// TIA Portal V21 export
DATA_BLOCK "Issue221_unitNested_readOnly"   // DB
{ S7_Optimized_Access := 'TRUE' }
// stored: AutoNumber true
BEGIN
END_DATA_BLOCK
